Fanuc KAREL source: KA00206.KL

PROGRAM KA00206
%NOLOCKGROUP
VAR
  SRC: ARRAY[4] OF VECTOR
  DST: ARRAY[4] OF XYZWPR
BEGIN
  DST = SRC
END KA00206
